Fanuc KAREL source: KD00076.KL

PROGRAM KD00076
%NOLOCKGROUP
VAR
  I: INTEGER
  J: INTEGER
  B: BOOLEAN
  R: REAL
  S: STRING[80]
BEGIN
  PURGE CONDITION[1]
END KD00076
